// CFC twin of T_SafeXor_Tests: the same tests drawn as CFC diagrams, the way a TwinSAFE project is authored.
    FUNCTION_BLOCK T_SafeXor_Tests_CFC EXTENDS T_SafeCfcTestSuite
    VAR
    // Test_ConnectedPairsAreExclusiveOr
    group_1 : T_SafeGroup;
    fb_1 : T_SafeXor(group := group_1);
END_VAR

Test_ConnectedPairsAreExclusiveOr();

METHOD PRIVATE Test_ConnectedPairsAreExclusiveOr
// note: this text did not pass the execution check against the stored diagram
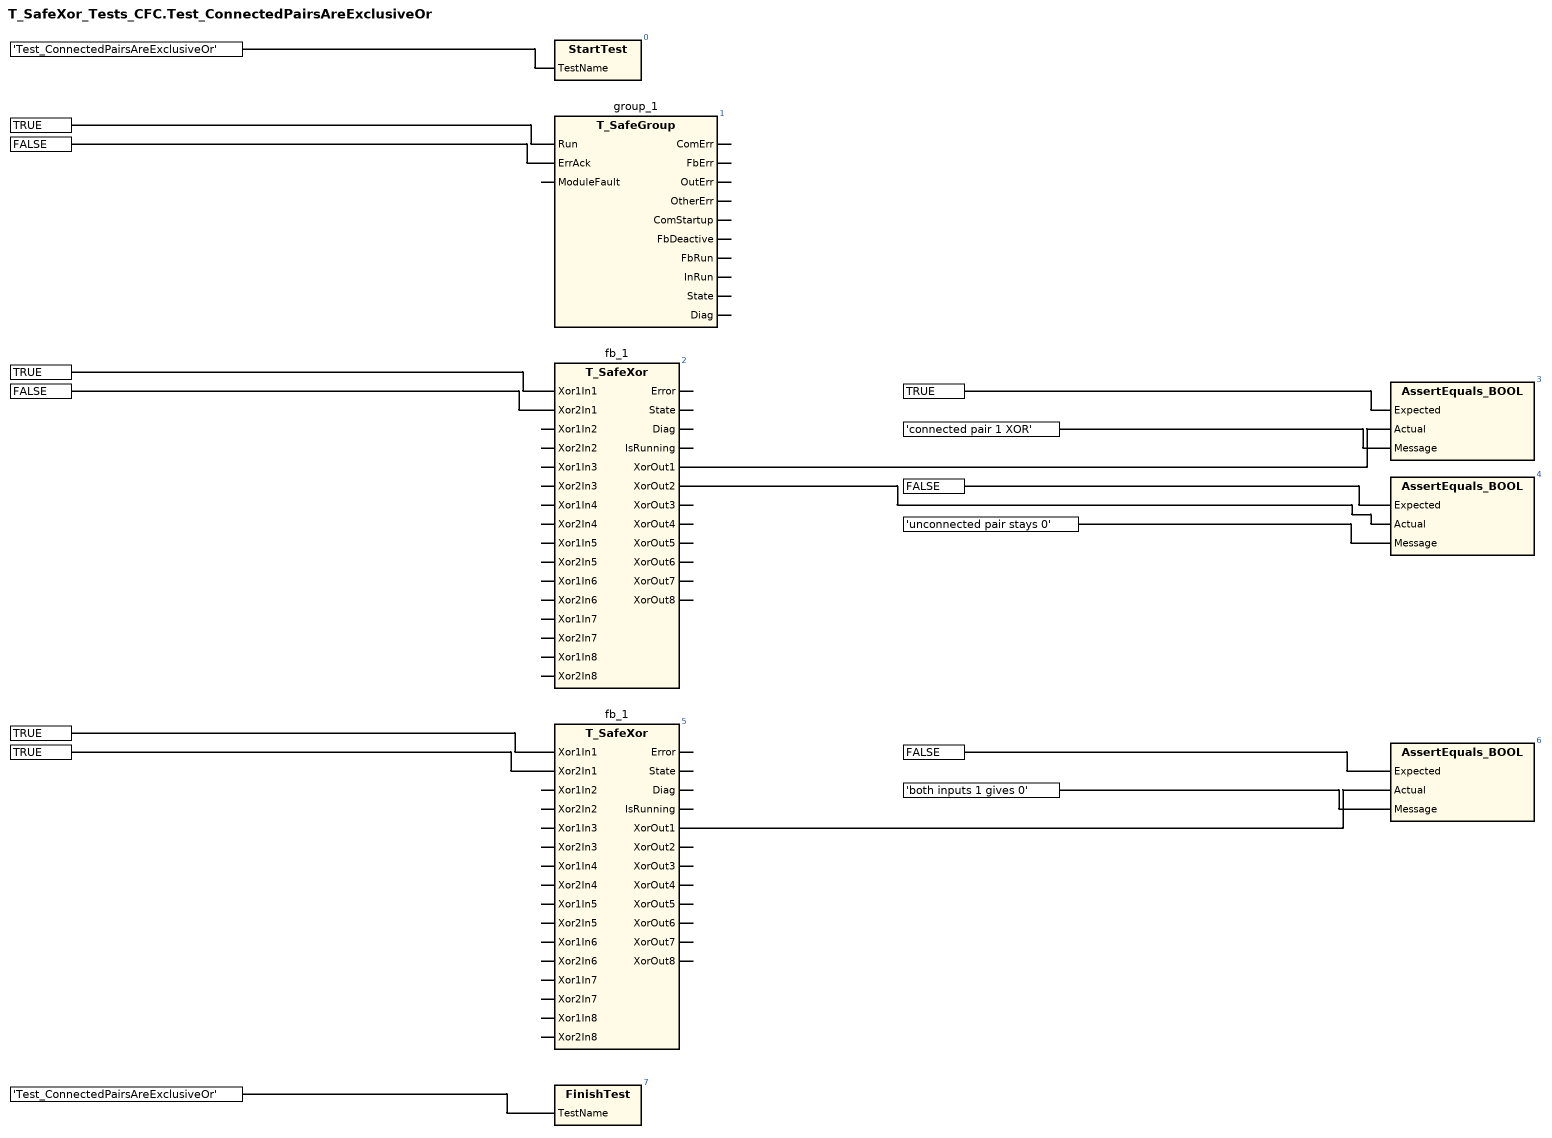
StartTest(TestName := 'Test_ConnectedPairsAreExclusiveOr');
group_1(Run := TRUE, ErrAck := FALSE); // T_SafeGroup
fb_1(Xor1In1 := TRUE, Xor2In1 := FALSE); // T_SafeXor
AssertEquals_BOOL(Expected := TRUE, Actual := fb_1.XorOut1, Message := 'connected pair 1 XOR');
AssertEquals_BOOL(Expected := FALSE, Actual := fb_1.XorOut2, Message := 'unconnected pair stays 0');
fb_1(Xor1In1 := TRUE, Xor2In1 := TRUE); // T_SafeXor
AssertEquals_BOOL(Expected := FALSE, Actual := fb_1.XorOut1, Message := 'both inputs 1 gives 0');
FinishTest(TestName := 'Test_ConnectedPairsAreExclusiveOr');
END_METHOD

END_FUNCTION_BLOCK

(* stored: Version 1.1.0.1, ProductVersion 3.1.4026.22
   POU T_SafeXor_Tests_CFC: Id {bf3107c6-cd29-5beb-a1b3-de80c7c3c5a0}, SpecialFunc None
   Method Test_ConnectedPairsAreExclusiveOr: Id {0de42657-bb8a-5a13-adbf-abfa96e22f52} *)
